(*
SPDX-FileCopyrightText: © 2026 Oleksandr Tiutyk <trofimich@gmail.com>
SPDX-License-Identifier: MIT
License: https://opensource.org/license/mit
*)

(*!
<summary>Runs one contract scenario and reports its own result.</summary>
<description>
Borrows the group fixture. The owning group serializes its cases in one task. AfterTest clears the fixture
after a successful run or an interrupted scenario. Terminal allocation failure uses the task boundary.
</description>
*)

{attribute 'no_assign'}
{attribute 'no_explicit_call' := 'do not call this function block directly'}
FUNCTION_BLOCK CollectionsContractTestCase EXTENDS TOF_Testing.SingleCycleTest
VAR_STAT
	{attribute 'hide'}
	_ClassName : STRING := __POUNAME();
END_VAR
VAR
	_Fixture : REFERENCE TO CollectionsContractTestFixture;
	_Scenario : COLLECTIONS_CONTRACT_SCENARIO;
END_VAR

(*!
<summary>Binds the group fixture and selects this case scenario.</summary>
<description>
Stores a borrowed reference without invoking the fixture. The owning group keeps it alive and
serializes use. TestElement initializes the name and parent.
</description>
<param name="name">Display name of this case.</param>
<param name="parent">Owning group.</param>
<param name="fixture">Live fixture owned by the group.</param>
<param name="scenario">Scenario assigned to this case.</param>
*)
METHOD FB_init : BOOL
VAR_INPUT
	bInitRetains: BOOL; // TRUE: the retain variables are initialized (reset warm / reset cold)
	bInCopyCode: BOOL; // TRUE: the instance will be copied to the copy code afterward (online change)
	name : WSTRING;
	parent : TOF_Testing.ITestElement;
	fixture : REFERENCE TO CollectionsContractTestFixture;
	scenario : COLLECTIONS_CONTRACT_SCENARIO;
END_VAR
IF NOT bInCopyCode THEN
	_Fixture REF= fixture;
	_Scenario := scenario;
END_IF

FB_init := TRUE;
END_METHOD

(*!
<summary>Runs the chosen scenario with the current assertions.</summary>
<description>
The fixture stays available to AfterTest if a call interrupts the scenario.
</description>
*)
METHOD PROTECTED ExecuteTest
VAR
	assertions : REFERENCE TO TOF_Testing.Assertions;
END_VAR
IF NOT __ISVALIDREF(_Fixture) THEN
	RecordFailure(message := "Missing collection contract fixture");

	RETURN;
END_IF

assertions REF= Assert;
_Fixture.ExecuteScenario(scenario := _Scenario, assertions := assertions);
END_METHOD

(*!
<summary>Clears the shared fixture and reports failed checked releases.</summary>
<description>
The fixture releases cursors before their sources. Cleanup preserves the first test failure and logs
any subsequent disposal failure.
</description>
*)
METHOD PROTECTED AfterTest
IF NOT __ISVALIDREF(_Fixture) THEN
	RETURN;
END_IF

IF NOT _Fixture.FinishScenario() THEN
	IF Outcome = TOF_Testing.TEST_OUTCOME.FAILED THEN
		Tc2_System.ADSLOGSTR(
			msgCtrlMask := Tc2_System.Global_Variables.ADSLOG_MSGTYPE_ERROR,
			msgFmtStr := 'Collection contract fixture cleanup failed in %s',
			strArg := TO_STRING(Name)
		);
	ELSE
		RecordFailure(message := "Collection contract fixture cleanup failed");
	END_IF
END_IF
END_METHOD

//! <summary>Borrows the concrete class name. Callers must not modify it.</summary>
{attribute 'monitoring' := 'call'}
PROPERTY ClassName : REFERENCE TO STRING
GET
ClassName REF= _ClassName;
END_GET
END_PROPERTY

//! <summary>Borrows the compiler-initialized namespace name. Callers must not modify it.</summary>
{attribute 'monitoring' := 'call'}
PROPERTY NamespaceName : REFERENCE TO STRING
GET
NamespaceName REF= CurrentNamespace.Name;
END_GET
END_PROPERTY

//! <summary>Reports the concrete instance size in bytes.</summary>
{attribute 'monitoring' := 'call'}
PROPERTY SelfSize : ULINT
GET
SelfSize := XSIZEOF(THIS^);
END_GET
END_PROPERTY

END_FUNCTION_BLOCK

(* stored: Version 1.1.0.1
   POU CollectionsContractTestCase: Id {09213e51-3db0-4f04-aaf0-6974e3d0b778}, SpecialFunc None
   Method FB_init: Id {6dcf16ce-b62f-4ce9-a6bc-617a87b0163b}
   Method ExecuteTest: Id {47d3479c-a695-4b8c-b216-509704468201}
   Method AfterTest: Id {8dcf536d-cd16-4e0e-bd03-ed16591b7f88}
   Property ClassName: Id {e331bb1c-f8d3-4996-9297-a6ba3ee1b0b5}
   Get Get: Id {e278a293-b085-49d5-acb3-16d4529832d3}
   Property NamespaceName: Id {bb5478b2-db99-4486-957e-938dce74a810}
   Get Get: Id {044ffc15-d6ea-4cb6-add6-e94baa6c70c7}
   Property SelfSize: Id {93c90dbe-316e-414c-8233-1662d41e079a}
   Get Get: Id {0b411ef9-461e-4216-a527-81a2d74a7392} *)
